(* IEC 61131-3 sources: hub-simuladores/simuladores/estacao-bombeamento-tq01/mastertool, 4 files *)

(* ---- GVL_SIM.st ---- *)
(* =====================================================================================
   GVL_SIM — Estação TQ-01 · CODESYS como servidor Modbus TCP (Modbus TCP Slave Device)
   Gerada da tabela "Variáveis e endereços" do simulador: as mesmas 22 variáveis, com o mesmo nome,
   tipo, endereço e significado. Cada uma está presa ao seu endereço com AT: não há programa de cópia.
   O comentário de cada variável é o texto da coluna "Significado" da tabela.

   Canal analógico como no hardware: LT01_Bruto é a contagem do A/D (0..32767 = 4..20 mA) e Ref_Bruto é a
   contagem do D/A (0..32767 = 0..10 V); o escalonamento é feito no seu programa.
   IHM: velocidade em % inteiro (75 = 75 %); setpoint e nível em centímetros (200 = 2,00 m).

   Configure o Modbus TCP Slave Device assim (aba de configuração):
       porta 502 · Unit ID 1 · Holding registers 4 · Input registers 3 · Coils 9 · Discrete inputs 6
   Com isso o CODESYS coloca, na aba "Modbus TCP Slave Device I/O Mapping":
       Holding Registers em %IW0 · Coils em %IB8 (%IX8.0…) · Input Registers em %QW0 · Discrete Inputs em %QB6 (%QX6.0…)
   Se algum endereço inicial for diferente no seu projeto, ajuste os AT abaixo (ou mude as quantidades acima).
   ===================================================================================== *)
VAR_GLOBAL
    (* ================= Simulador → CLP (o simulador escreve, o CLP lê) ================= *)
    S1_Liga        AT %IX8.0  : BOOL;   (* Botoeira S1 liga (NA): 1 enquanto pressionada *)
    S2_Desliga_NF  AT %IX8.1  : BOOL;   (* Botoeira S2 desliga (NF): 1 em repouso, 0 pressionada *)
    S3_Reset       AT %IX8.2  : BOOL;   (* Botoeira S3 reset (NA) *)
    S4_Auto        AT %IX8.3  : BOOL;   (* Seletor S4: 1 = automático, 0 = manual *)
    S0_Emerg_NF    AT %IX8.4  : BOOL;   (* Emergência S0 (NF): 1 destravado, 0 acionado *)
    Inv_Rodando    AT %IX8.5  : BOOL;   (* Relé DO2 do CFW500 (F > Fx): inversor acima de 3 Hz *)
    Inv_OK         AT %IX8.6  : BOOL;   (* Relé DO1 do CFW500 (sem falha): 0 = falha ou sem alimentação *)
    LSHH           AT %IX8.7  : BOOL;   (* Chave de nível muito alto LSHH-01 (2,8 m) *)
    LSLL           AT %IX9.0  : BOOL;   (* Chave de nível muito baixo LSLL-01 (0,3 m) *)
    LT01_Bruto     AT %IW0    : INT;    (* Nível LT-01, contagem do A/D: 0–32767 = 4–20 mA = 0–3,5 m (negativo abaixo de 4 mA) *)
    HB_Sim         AT %IW1    : UINT;   (* Heartbeat do simulador: +1 por segundo *)
    IHM_Velocidade AT %IW2    : INT;    (* IHM: velocidade da bomba pedida pelo operador, em % (0–100) *)
    IHM_Setpoint   AT %IW3    : INT;    (* IHM: setpoint de nível para o automático, em cm (0–300; 200 = 2,00 m) *)

    (* ================= CLP → simulador (o CLP escreve, o simulador lê) ================= *)
    H1             AT %QX6.0  : BOOL;   (* Sinaleiro verde — em operação *)
    H2             AT %QX6.1  : BOOL;   (* Sinaleiro amarelo — alarme *)
    H3             AT %QX6.2  : BOOL;   (* Sinaleiro vermelho — falha *)
    H4             AT %QX6.3  : BOOL;   (* Sirene *)
    Inv_Gira       AT %QX6.4  : BOOL;   (* DI1 do CFW500: gira/para (em série com o 2º NF do S0) *)
    Inv_Reset      AT %QX6.5  : BOOL;   (* DI3 do CFW500: reset de falha (borda de subida) *)
    Ref_Bruto      AT %QW0    : INT;    (* Referência de velocidade, contagem do D/A: 0–32767 = 0–10 V = 0–60 Hz *)
    HB_CLP         AT %QW1    : UINT;   (* Heartbeat do CLP: +1 a cada 0,5 s *)
    IHM_Nivel      AT %QW2    : INT;    (* Nível que o CLP manda a IHM mostrar, em cm (152 = 1,52 m) *)
END_VAR

(* ---- GVL_SIMULADOR.st ---- *)
(* =====================================================================================
   GVL_SIMULADOR — Estação TQ-01 · CODESYS como servidor Modbus TCP (Modbus TCP Slave Device)
   Gerada da tabela "Variáveis e endereços" do simulador: as mesmas 22 variáveis, com o mesmo nome,
   tipo, endereço e significado. SEM AT: ligue cada uma ao seu canal pela coluna "Variable" da aba de mapeamento
   (botão "...", Application.GVL_SIMULADOR.<nome>). Não use AT junto com o mapeamento.
   O comentário de cada variável é o texto da coluna "Significado" da tabela.

   Canal analógico como no hardware: LT01_Bruto é a contagem do A/D (0..32767 = 4..20 mA) e Ref_Bruto é a
   contagem do D/A (0..32767 = 0..10 V); o escalonamento é feito no seu programa.
   IHM: velocidade em % inteiro (75 = 75 %); setpoint e nível em centímetros (200 = 2,00 m).

   Configure o Modbus TCP Slave Device assim (aba de configuração):
       porta 502 · Unit ID 1 · Holding registers 4 · Input registers 3 · Coils 9 · Discrete inputs 6
   Com isso o CODESYS coloca, na aba "Modbus TCP Slave Device I/O Mapping":
       Holding Registers em %IW0 · Coils em %IB8 (%IX8.0…) · Input Registers em %QW0 · Discrete Inputs em %QB6 (%QX6.0…)
   Se algum endereço inicial for diferente no seu projeto, ajuste os AT abaixo (ou mude as quantidades acima).
   ===================================================================================== *)
VAR_GLOBAL
    (* ================= Simulador → CLP (o simulador escreve, o CLP lê) ================= *)
    S1_Liga                   : BOOL;   (* Botoeira S1 liga (NA): 1 enquanto pressionada *)
    S2_Desliga_NF             : BOOL;   (* Botoeira S2 desliga (NF): 1 em repouso, 0 pressionada *)
    S3_Reset                  : BOOL;   (* Botoeira S3 reset (NA) *)
    S4_Auto                   : BOOL;   (* Seletor S4: 1 = automático, 0 = manual *)
    S0_Emerg_NF               : BOOL;   (* Emergência S0 (NF): 1 destravado, 0 acionado *)
    Inv_Rodando               : BOOL;   (* Relé DO2 do CFW500 (F > Fx): inversor acima de 3 Hz *)
    Inv_OK                    : BOOL;   (* Relé DO1 do CFW500 (sem falha): 0 = falha ou sem alimentação *)
    LSHH                      : BOOL;   (* Chave de nível muito alto LSHH-01 (2,8 m) *)
    LSLL                      : BOOL;   (* Chave de nível muito baixo LSLL-01 (0,3 m) *)
    LT01_Bruto                : INT;    (* Nível LT-01, contagem do A/D: 0–32767 = 4–20 mA = 0–3,5 m (negativo abaixo de 4 mA) *)
    HB_Sim                    : UINT;   (* Heartbeat do simulador: +1 por segundo *)
    IHM_Velocidade            : INT;    (* IHM: velocidade da bomba pedida pelo operador, em % (0–100) *)
    IHM_Setpoint              : INT;    (* IHM: setpoint de nível para o automático, em cm (0–300; 200 = 2,00 m) *)

    (* ================= CLP → simulador (o CLP escreve, o simulador lê) ================= *)
    H1                        : BOOL;   (* Sinaleiro verde — em operação *)
    H2                        : BOOL;   (* Sinaleiro amarelo — alarme *)
    H3                        : BOOL;   (* Sinaleiro vermelho — falha *)
    H4                        : BOOL;   (* Sirene *)
    Inv_Gira                  : BOOL;   (* DI1 do CFW500: gira/para (em série com o 2º NF do S0) *)
    Inv_Reset                 : BOOL;   (* DI3 do CFW500: reset de falha (borda de subida) *)
    Ref_Bruto                 : INT;    (* Referência de velocidade, contagem do D/A: 0–32767 = 0–10 V = 0–60 Hz *)
    HB_CLP                    : UINT;   (* Heartbeat do CLP: +1 a cada 0,5 s *)
    IHM_Nivel                 : INT;    (* Nível que o CLP manda a IHM mostrar, em cm (152 = 1,52 m) *)
    (* ================= Variáveis internas do CLP (não vão para a rede) ================= *)
    IHM_Nivel_Real            : REAL;   (* Nível do tanque em metros (IHM_Nivel / 100) *)
    IHM_Nivel_SP_Real         : REAL;   (* Nível que o operador envia através da IHM, neste caso já convertido *)
    IHM_Nivel_SP_Liga         : REAL;   (* Liga a bomba abaixo deste nível (SP − histerese) *)
    IHM_Nivel_SP_Desl         : REAL;   (* Desliga a bomba acima deste nível (SP + histerese) *)
END_VAR

(* ---- PRG_TQ01.st ---- *)
(* =====================================================================================
   PRG_TQ01 — bomba B-01 com intertravamentos, escalonamento do canal analógico de entrada (LT-01)
   e de saída (referência do inversor), IHM e heartbeat. Usa só os nomes da tabela (GVL_SIM).
   Chame na MainTask.
   Canal analógico como no hardware:
     entrada  LT01_Bruto : 0..32767 = 4..20 mA = 0..3,5 m   (negativo abaixo de 4 mA)
     saída    Ref_Bruto  : 0..32767 = 0..10 V  = 0..60 Hz
   IHM: IHM_Velocidade em % (0–100), IHM_Setpoint e IHM_Nivel em cm (200 = 2,00 m).
   Manual: a bomba roda na velocidade pedida na IHM.
   Automático: liga a 75 % abaixo de (setpoint − 0,5 m) e para acima de (setpoint + 0,5 m).
   ===================================================================================== *)
PROGRAM PRG_TQ01
VAR
    rNivel      : REAL;    (* nível do tanque em metros (escalonado do LT01_Bruto) *)
    rVelIHM     : REAL;    (* velocidade pedida na IHM, % *)
    rSetpoint   : REAL;    (* setpoint de nível da IHM, m *)
    rRefPct     : REAL;    (* referência que vai para o inversor, % *)
    rtLiga      : R_TRIG;
    xLigado     : BOOL;
    xFalha      : BOOL;
    xCondicao   : BOOL;
    xEnche      : BOOL;
    xFioRompido : BOOL;
    tonSimFora  : TON;
    uiHBAnt     : UINT;
    tonHB       : TON;
END_VAR

(* 1. Entrada analógica: escalonamento da contagem do A/D para metros *)
rNivel      := INT_TO_REAL(GVL_SIM.LT01_Bruto) / 32767.0 * 3.5;   (* 0..32767 = 0..3,5 m *)
xFioRompido := GVL_SIM.LT01_Bruto < -410;                          (* abaixo de 3,8 mA *)

(* IHM: velocidade já vem em %; setpoint vem em cm *)
rVelIHM   := LIMIT(0.0, INT_TO_REAL(GVL_SIM.IHM_Velocidade), 100.0);
rSetpoint := LIMIT(0.0, INT_TO_REAL(GVL_SIM.IHM_Setpoint) / 100.0, 3.0);      (* cm -> m *)

(* 2. Watchdog: HB_Sim parado por 3 s = simulador fora *)
tonSimFora(IN := (GVL_SIM.HB_Sim = uiHBAnt), PT := T#3S);
uiHBAnt := GVL_SIM.HB_Sim;

(* 3. Intertravamentos (S2 e S0 são NF: 1 em repouso) *)
xCondicao := GVL_SIM.S2_Desliga_NF AND GVL_SIM.S0_Emerg_NF AND GVL_SIM.Inv_OK
         AND NOT GVL_SIM.LSHH AND NOT xFioRompido AND NOT tonSimFora.Q;

IF GVL_SIM.S3_Reset THEN
    xFalha := FALSE;
END_IF
IF NOT xCondicao THEN
    IF xLigado THEN
        xFalha := TRUE;
    END_IF
    xLigado := FALSE;
END_IF
rtLiga(CLK := GVL_SIM.S1_Liga);
IF rtLiga.Q AND xCondicao AND NOT xFalha THEN
    xLigado := TRUE;
END_IF

(* 4. Manual x automático *)
IF GVL_SIM.S4_Auto THEN
    IF rNivel < rSetpoint - 0.5 THEN
        xEnche := TRUE;
    ELSIF rNivel > rSetpoint + 0.5 THEN
        xEnche := FALSE;
    END_IF
    GVL_SIM.Inv_Gira := xLigado AND xEnche;
    rRefPct := 75.0;
ELSE
    xEnche := FALSE;
    GVL_SIM.Inv_Gira := xLigado;
    rRefPct := rVelIHM;
END_IF
IF NOT GVL_SIM.Inv_Gira THEN
    rRefPct := 0.0;
END_IF

(* 5. Saída analógica: escalonamento de % para a contagem do D/A (0..32767 = 0..10 V) *)
GVL_SIM.Ref_Bruto := REAL_TO_INT(rRefPct / 100.0 * 32767.0);

(* 6. Sinalização, reset do inversor e IHM *)
GVL_SIM.H1 := GVL_SIM.Inv_Rodando;
GVL_SIM.H2 := rNivel > 2.6 OR rNivel < 0.5 OR GVL_SIM.LSHH OR GVL_SIM.LSLL;
GVL_SIM.H3 := xFalha;
GVL_SIM.H4 := xFalha AND NOT GVL_SIM.S3_Reset;
GVL_SIM.Inv_Reset := GVL_SIM.S3_Reset;
GVL_SIM.IHM_Nivel := REAL_TO_INT(rNivel * 100.0);                (* m -> cm *)

(* 7. Heartbeat do CLP: +1 a cada 500 ms *)
tonHB(IN := NOT tonHB.Q, PT := T#500MS);
IF tonHB.Q THEN
    GVL_SIM.HB_CLP := GVL_SIM.HB_CLP + 1;
END_IF

(* ---- PRG_TQ01_GVL_SIMULADOR.st ---- *)
(* =====================================================================================
   PRG_TQ01 — Estação TQ-01, com a GVL_SIMULADOR. Equivale ao programa em Ladder da aula:
     · cálculos do canal analógico e da IHM (ST)
     · automático liga-desliga com HISTERESE de ± 10 cm, sem TON:
         liga  (SET)   quando IHM_Nivel_Real <= IHM_Nivel_SP_Liga  (SP − 0,10 m)
         desliga (RESET) quando IHM_Nivel_Real >= IHM_Nivel_SP_Desl (SP + 0,10 m)
         entre os dois, Inv_Gira fica como está
     · degrau de segurança: sai do automático, emergência ou LSHH -> RESET do Inv_Gira
   A velocidade da bomba é sempre a pedida na IHM (IHM_Velocidade).
   ===================================================================================== *)
PROGRAM PRG_TQ01
VAR
    tonHB : TON;    (* heartbeat do CLP *)
END_VAR

(* ---------- cálculos (canal analógico e IHM) ---------- *)
GVL_SIMULADOR.Ref_Bruto         := REAL_TO_INT(GVL_SIMULADOR.IHM_Velocidade / 100.0 * 32767.0);   (* % -> contagem do D/A *)
GVL_SIMULADOR.IHM_Nivel         := REAL_TO_INT((GVL_SIMULADOR.LT01_Bruto) / 32767.0 * 350);       (* contagem do A/D -> cm *)
GVL_SIMULADOR.IHM_Nivel_Real    := TO_REAL(GVL_SIMULADOR.IHM_Nivel) / 100.0;                      (* cm -> m *)
GVL_SIMULADOR.IHM_Nivel_SP_Real := LIMIT(0.5, INT_TO_REAL(GVL_SIMULADOR.IHM_Setpoint) / 100.0, 2.6); (* cm -> m, SP entre 0,5 e 2,6 m *)
GVL_SIMULADOR.IHM_Nivel_SP_Liga := GVL_SIMULADOR.IHM_Nivel_SP_Real - 0.10;                        (* histerese: liga 10 cm abaixo *)
GVL_SIMULADOR.IHM_Nivel_SP_Desl := GVL_SIMULADOR.IHM_Nivel_SP_Real + 0.10;                        (* histerese: desliga 10 cm acima *)

(* ---------- degrau 1: automático — liga (SET) ---------- *)
IF GVL_SIMULADOR.S4_Auto AND GVL_SIMULADOR.S0_Emerg_NF AND NOT GVL_SIMULADOR.LSHH
   AND GVL_SIMULADOR.IHM_Nivel_Real <= GVL_SIMULADOR.IHM_Nivel_SP_Liga THEN
    GVL_SIMULADOR.Inv_Gira := TRUE;
END_IF

(* ---------- degrau 2: automático — desliga (RESET) ---------- *)
IF GVL_SIMULADOR.S4_Auto AND GVL_SIMULADOR.S0_Emerg_NF AND NOT GVL_SIMULADOR.LSHH
   AND GVL_SIMULADOR.IHM_Nivel_Real >= GVL_SIMULADOR.IHM_Nivel_SP_Desl THEN
    GVL_SIMULADOR.Inv_Gira := FALSE;
END_IF

(* ---------- degrau 3: segurança — sai do automático, emergência ou LSHH (RESET) ---------- *)
IF NOT GVL_SIMULADOR.S4_Auto OR NOT GVL_SIMULADOR.S0_Emerg_NF OR GVL_SIMULADOR.LSHH THEN
    GVL_SIMULADOR.Inv_Gira := FALSE;
END_IF

(* ---------- sinalização e reset do inversor ---------- *)
GVL_SIMULADOR.H1 := GVL_SIMULADOR.Inv_Rodando;
GVL_SIMULADOR.H2 := GVL_SIMULADOR.LSHH OR GVL_SIMULADOR.LSLL;
GVL_SIMULADOR.H3 := NOT GVL_SIMULADOR.Inv_OK;
GVL_SIMULADOR.Inv_Reset := GVL_SIMULADOR.S3_Reset;

(* ---------- heartbeat do CLP: +1 a cada 500 ms ---------- *)
tonHB(IN := NOT tonHB.Q, PT := T#500MS);
IF tonHB.Q THEN
    GVL_SIMULADOR.HB_CLP := GVL_SIMULADOR.HB_CLP + 1;
END_IF
